FUNCTION_BLOCK FB_IoInput IMPLEMENTS I_IoBit;

VAR
	
	_bHw	AT %I* : BOOL;
	_ftrig			: F_TRIG;
	_rtrig			: R_TRIG;
	_Q				: BOOL;
END_VAR

_Q		:= _bHw;

_rtrig( CLK := _bHw );
_ftrig( CLK := _bHw );

//FB_Init is always available implicitly and it is used primarily for initialization.
//The return value is not evaluated. For a specific influence, you can also declare the
//methods explicitly and provide additional code there with the standard initialization
//code. You can evaluate the return value.
METHOD FB_Init: BOOL
VAR_INPUT
    bInitRetains: BOOL; // TRUE: the retain variables are initialized (reset warm / reset cold)
    bInCopyCode: BOOL;  // TRUE: the instance will be copied to the copy code afterward (online change)
	IoGroup		: I_IoGroup;   
END_VAR
IoGroup.AddIo(THIS^);
END_METHOD


PROPERTY ftrig : BOOL
GET
ftrig := _ftrig.Q;
END_GET
SET
END_SET
END_PROPERTY

PROPERTY Q : BOOL
GET
Q := _Q;
END_GET
SET
END_SET
END_PROPERTY


PROPERTY rtrig : BOOL
GET
rtrig := _rtrig.Q;
END_GET
SET
END_SET
END_PROPERTY


METHOD Update
THIS^();
END_METHOD

END_FUNCTION_BLOCK

(* stored: Version 1.1.0.1
   POU FB_IoInput: Id {2798f21f-b023-4222-b3a7-e9218e155a00}, SpecialFunc None
   Method FB_Init: Id {c6a4cc9b-1c14-4c14-a1aa-8ace61b447fd}
   Property ftrig: Id {30053e0b-3ef4-4010-bcf9-40deb03c8b04}
   Get Get: Id {131e45ce-1000-4ca9-adb8-dd46c6b76458}
   Set Set: Id {44bfd57b-aa6d-4431-892e-bf440952ab25}
   Property Q: Id {6f3b9111-930a-41c9-b977-552d568d2f92}
   Get Get: Id {485dc2d8-603c-4cdd-b225-0e52a16edfd6}
   Set Set: Id {a4b3e9ca-f778-48e5-94bf-036304326822}
   Property rtrig: Id {f2c14d3c-edf5-469c-acd3-dcb4ab0b8ef9}
   Get Get: Id {6f8b5bdf-30ae-46ad-b9f4-843888573183}
   Set Set: Id {ba2e0ca5-cff0-49e2-a84e-f88fc1a91f85}
   Method Update: Id {a3b0ff73-c1c7-4cf3-baa1-8ef4b5b9f3ba} *)
